FUNCTION_BLOCK IDENTIFICATION_UPDATE_GATE (* Experimental; offline checks only; native export/runtime pending *)
  (* Standard: 61499-2 *)
  (* Version 0.1, 2026-10-20, Guilherme *)
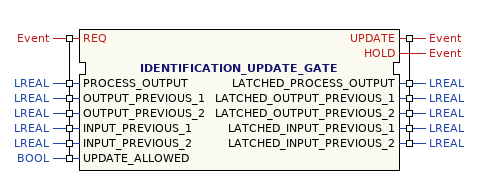
  EVENT_INPUT
    REQ WITH PROCESS_OUTPUT, OUTPUT_PREVIOUS_1, OUTPUT_PREVIOUS_2, INPUT_PREVIOUS_1, INPUT_PREVIOUS_2, UPDATE_ALLOWED;
  END_EVENT
  EVENT_OUTPUT
    UPDATE WITH LATCHED_PROCESS_OUTPUT, LATCHED_OUTPUT_PREVIOUS_1, LATCHED_OUTPUT_PREVIOUS_2, LATCHED_INPUT_PREVIOUS_1, LATCHED_INPUT_PREVIOUS_2;
    HOLD;
  END_EVENT
  VAR_INPUT
    PROCESS_OUTPUT : LREAL;
    OUTPUT_PREVIOUS_1 : LREAL;
    OUTPUT_PREVIOUS_2 : LREAL;
    INPUT_PREVIOUS_1 : LREAL;
    INPUT_PREVIOUS_2 : LREAL;
    UPDATE_ALLOWED : BOOL;
  END_VAR
  VAR_OUTPUT
    LATCHED_PROCESS_OUTPUT : LREAL;
    LATCHED_OUTPUT_PREVIOUS_1 : LREAL;
    LATCHED_OUTPUT_PREVIOUS_2 : LREAL;
    LATCHED_INPUT_PREVIOUS_1 : LREAL;
    LATCHED_INPUT_PREVIOUS_2 : LREAL;
  END_VAR
  VAR
    ALLOW_CAPTURED : BOOL;
  END_VAR
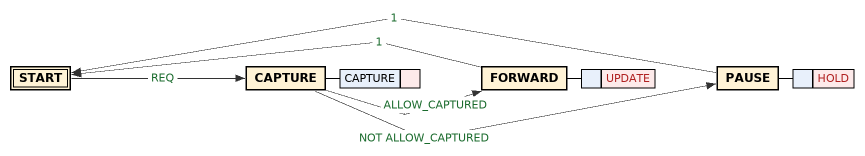
  EC_STATES
    START;
    CAPTURE : CAPTURE;
    FORWARD : -> UPDATE;
    PAUSE : -> HOLD;
  END_STATES
  EC_TRANSITIONS
    START TO CAPTURE := REQ;
    CAPTURE TO FORWARD := ALLOW_CAPTURED;
    CAPTURE TO PAUSE := NOT ALLOW_CAPTURED;
    FORWARD TO START := 1;
    PAUSE TO START := 1;
  END_TRANSITIONS
  ALGORITHM CAPTURE IN ST:
ALLOW_CAPTURED := UPDATE_ALLOWED;
IF ALLOW_CAPTURED THEN
LATCHED_PROCESS_OUTPUT := PROCESS_OUTPUT;
LATCHED_OUTPUT_PREVIOUS_1 := OUTPUT_PREVIOUS_1;
LATCHED_OUTPUT_PREVIOUS_2 := OUTPUT_PREVIOUS_2;
LATCHED_INPUT_PREVIOUS_1 := INPUT_PREVIOUS_1;
LATCHED_INPUT_PREVIOUS_2 := INPUT_PREVIOUS_2;
END_IF;
  END_ALGORITHM
END_FUNCTION_BLOCK
